(*
This is a paragraph.

Paragraphs line up at their left edges, and are normally separated 
by blank lines.
*)

FUNCTION_BLOCK FB_Libdoc_Paragraph
VAR_INPUT
    nVarA : INT;
    nVarB : INT;
END_VAR
VAR_OUTPUT
    nSum : INT;
END_VAR
VAR
END_VAR

END_FUNCTION_BLOCK

(* stored: Version 1.1.0.1, ProductVersion 3.1.4022.18
   POU FB_Libdoc_Paragraph: Id {53c81225-e4bc-429a-8ffd-21458727dad8}, SpecialFunc None *)
